Staubli VAL3: selStartUpProg.pgx

public program selStartUpProg()
begin
  nProgType=1
end
